(* PLC project PR_TT-1MasterSeq_Soft2.0_workflow_b380e4_PLC, SiemensToBackhoff Siemens TIA Portal → Beckhoff TwinCAT PLCopen Converter 2.2 *)
(* stored: creationDateTime 2026-10-12T09:25:48.748496, modificationDateTime 2026-10-12T09:25:48.748496 *)

FUNCTION_BLOCK PR_TT-1MasterSeq_Soft2.0_workflow_b380e4
VAR_INPUT
	iAllStationProcessOver : BOOL;
	iAutoRunning : BOOL;
	iHiPotTestOver_1 : BOOL;
	iHiPotTestOver_2 : BOOL;
	iHiPot_RTR_1 : BOOL;
	iHiPot_RTR_2 : BOOL;
	iIndexOver : BOOL;
	iIndex_RTR_Place1 : BOOL;
	iIndex_RTR_Place2 : BOOL;
	iOTS_Frm_Shuttle_1 : BOOL;
	iOTS_Frm_Shuttle_2 : BOOL;
	iOTS_Frm_TransferGantry : BOOL;
	iOperatorAck : BOOL;
	iPartPickOver : BOOL;
	iPartPickOver_1 : BOOL;
	iPartPickOver_2 : BOOL;
	iPartPlaceByTransferGantry : BOOL;
	iPartPlaceOver_IFGantry : BOOL;
	iPartPlaceOver_IndexPlace1 : BOOL;
	iPartPlaceOver_IndexPlace2 : BOOL;
	iPartPresent_IFGantry : BOOL;
	iPartPresent_Shuttle_1 : BOOL;
	iPartPresent_Shuttle_2 : BOOL;
	iPartPresent_TxGantry_1 : BOOL;
	iPartPresent_TxGantry_2 : BOOL;
	iRTR_Frm_TransferGantry_1 : BOOL;
	iRTR_Frm_TransferGantry_2 : BOOL;
	iReset_fault : BOOL;
	iShuttleReadyToReceive : BOOL;
	iSstMode : BOOL;
	iSstPB : BOOL;
END_VAR
VAR_OUTPUT
	qError : ARRAY[1..1] OF BOOL;
	qInfeedGantry_PickStart : BOOL;
	qInfeedGantry_PlaceStart : BOOL;
	qShuttle_1PickStart : BOOL;
	qShuttle_1PlaceStart : BOOL;
	qShuttle_2PickStart : BOOL;
	qShuttle_2PlaceStart : BOOL;
	qTransferGantry1_PickStart : BOOL;
	qTransferGantry1_PlaceStart : BOOL;
	qTransferGantry2_PickStart : BOOL;
	qTransferGantry2_PlaceStart : BOOL;
END_VAR
VAR
	c10_ChkPartStsAtSubStn_T1 : BOOL;
	c10_ChkPartStsAtSubStn_T2 : BOOL;
	c10_ChkPartStsAtSubStn_T3 : BOOL;
	c10_ChkPartStsAtSubStn_T4 : BOOL;
	c10_ChkPartStsAtSubStn_T5 : BOOL;
	c10_ChkPartStsAtSubStn_T6 : BOOL;
	c10_ChkPartStsAtSubStn_T7 : BOOL;
	c130_ChkPartPrsntStsShuttle2_T1 : BOOL;
	c130_ChkPartPrsntStsShuttle2_T2 : BOOL;
	c200_ChkPartPrsntTxGantry1_T1 : BOOL;
	c200_ChkPartPrsntTxGantry1_T2 : BOOL;
	c250_ChkPartPrsntTxGantry2_T1 : BOOL;
	c250_ChkPartPrsntTxGantry2_T2 : BOOL;
	c300_ChkPartPrsntIndexer_T1 : BOOL;
	c300_ChkPartPrsntIndexer_T2 : BOOL;
	c30_ChkPartStsIFGantry_T1 : BOOL;
	c30_ChkPartStsIFGantry_T2 : BOOL;
	c70_ChkPartPrsntStsShuttle1_T1 : BOOL;
	c70_ChkPartPrsntStsShuttle1_T2 : BOOL;
	StateNo : INT;
	s100_WtHiPotTestOver1 : BOOL;
	s100_WtHiPotTestOver1_T1 : BOOL;
	s10_ChkPartStsAtSubStn : BOOL;
	s10_ChkPartStsAtSubStn_T1 : BOOL;
	s10_ChkPartStsAtSubStn_T2 : BOOL;
	s10_ChkPartStsAtSubStn_T3 : BOOL;
	s10_ChkPartStsAtSubStn_T4 : BOOL;
	s10_ChkPartStsAtSubStn_T5 : BOOL;
	s10_ChkPartStsAtSubStn_T6 : BOOL;
	s10_ChkPartStsAtSubStn_T7 : BOOL;
	s110_WtTxGantryRTR1 : BOOL;
	s110_WtTxGantryRTR1_T1 : BOOL;
	s120_WtPartUnldOvrTxGantry1 : BOOL;
	s120_WtPartUnldOvrTxGantry1_T1 : BOOL;
	s130_ChkPartPrsntStsShuttle2 : BOOL;
	s130_ChkPartPrsntStsShuttle2_T1 : BOOL;
	s130_ChkPartPrsntStsShuttle2_T2 : BOOL;
	s140_WtIFGantryPlacePart2 : BOOL;
	s140_WtIFGantryPlacePart2_T1 : BOOL;
	s150_WtHiPotRdyRcvPart2 : BOOL;
	s150_WtHiPotRdyRcvPart2_T1 : BOOL;
	s160_WtHiPotTestOver2 : BOOL;
	s160_WtHiPotTestOver2_T1 : BOOL;
	s170_WtTxGantryRTR2 : BOOL;
	s170_WtTxGantryRTR2_T1 : BOOL;
	s190_WtPartUnldOvrTxGantry2 : BOOL;
	s190_WtPartUnldOvrTxGantry2_T1 : BOOL;
	s1_WtResetRel : BOOL;
	s1_WtResetRel_T1 : BOOL;
	s200_ChkPartPrsntTxGantry1 : BOOL;
	s200_ChkPartPrsntTxGantry1_T1 : BOOL;
	s200_ChkPartPrsntTxGantry1_T2 : BOOL;
	s20_WtOperatorAck : BOOL;
	s20_WtOperatorAck_T1 : BOOL;
	s210_WtShuttle1RdySendPal : BOOL;
	s210_WtShuttle1RdySendPal_T1 : BOOL;
	s220_WtPartPickTxGantry1 : BOOL;
	s220_WtPartPickTxGantry1_T1 : BOOL;
	s230_WtIndexRTRPlace1 : BOOL;
	s230_WtIndexRTRPlace1_T1 : BOOL;
	s240_WtPartPlaceOverIndexPlace1 : BOOL;
	s240_WtPartPlaceOverIndexPlace1_T1 : BOOL;
	s250_ChkPartPrsntTxGantry2 : BOOL;
	s250_ChkPartPrsntTxGantry2_T1 : BOOL;
	s250_ChkPartPrsntTxGantry2_T2 : BOOL;
	s260_WtShuttle2RdySendPal : BOOL;
	s260_WtShuttle2RdySendPal_T1 : BOOL;
	s270_WtPartPickTxGantry2 : BOOL;
	s270_WtPartPickTxGantry2_T1 : BOOL;
	s280_WtIndexRTRPlace2 : BOOL;
	s280_WtIndexRTRPlace2_T1 : BOOL;
	s290_WtPartPlaceOverIndexPlace2 : BOOL;
	s290_WtPartPlaceOverIndexPlace2_T1 : BOOL;
	s300_ChkPartPrsntIndexer : BOOL;
	s300_ChkPartPrsntIndexer_T1 : BOOL;
	s300_ChkPartPrsntIndexer_T2 : BOOL;
	s30_ChkPartStsIFGantry : BOOL;
	s30_ChkPartStsIFGantry_T1 : BOOL;
	s30_ChkPartStsIFGantry_T2 : BOOL;
	s310_WtOTSFrmTxGantry : BOOL;
	s310_WtOTSFrmTxGantry_T1 : BOOL;
	s320_WtPartPlaceByTxGantry : BOOL;
	s320_WtPartPlaceByTxGantry_T1 : BOOL;
	s330_WtAllStnProcessOver : BOOL;
	s330_WtAllStnProcessOver_T1 : BOOL;
	s340_WtIndexOver : BOOL;
	s340_WtIndexOver_T1 : BOOL;
	s40_WtPartPickOverIFGantry : BOOL;
	s40_WtPartPickOverIFGantry_T1 : BOOL;
	s50_WtShuttleRdyRcvPart : BOOL;
	s50_WtShuttleRdyRcvPart_T1 : BOOL;
	s60_WtPartPlaceByGantry : BOOL;
	s60_WtPartPlaceByGantry_T1 : BOOL;
	s70_ChkPartPrsntStsShuttle1 : BOOL;
	s70_ChkPartPrsntStsShuttle1_T1 : BOOL;
	s70_ChkPartPrsntStsShuttle1_T2 : BOOL;
	s80_WtIFGantryPlacePart : BOOL;
	s80_WtIFGantryPlacePart_T1 : BOOL;
	s90_WtHiPotRdyRcvPart1 : BOOL;
	s90_WtHiPotRdyRcvPart1_T1 : BOOL;
	sAbnormalCondition : BOOL;
	sIndexerSeq : BOOL;
	sInfeedGantry : BOOL;
	sPartAbsentAtAllStn : BOOL;
	sPartPrsntAtStn : BOOL;
	sShuttle_1Seq : BOOL;
	sShuttle_2Seq : BOOL;
	sSst : BOOL;
	sSstPulse : BOOL;
	sSstRise : R_TRIG;
	sStWtResetRel : BOOL;
	sStWtResetRel_T1 : BOOL;
	sTransferGantry_1Seq : BOOL;
	sTransferGantry_2Seq : BOOL;
END_VAR
VAR_TEMP
	tOne : BOOL;
END_VAR
  VAR  (* added by the conversion: wires and edge detectors of the diagram *)
    _w24 : BOOL;
    _w26 : BOOL;
    _w39 : BOOL;
    _w41 : BOOL;
    _w42 : BOOL;
    _w116 : BOOL;
    _w119 : BOOL;
    _w120 : BOOL;
    _w121 : BOOL;
    _w122 : BOOL;
    _w123 : BOOL;
    _w124 : BOOL;
    _w125 : BOOL;
    _w126 : BOOL;
    _w139 : BOOL;
    _w141 : BOOL;
    _w142 : BOOL;
    _w170 : BOOL;
    _w174 : BOOL;
    _w175 : BOOL;
    _w176 : BOOL;
    _w190 : BOOL;
    _w192 : BOOL;
    _w193 : BOOL;
    _w210 : BOOL;
    _w212 : BOOL;
    _w213 : BOOL;
    _w226 : BOOL;
    _w228 : BOOL;
    _w229 : BOOL;
    _w257 : BOOL;
    _w261 : BOOL;
    _w262 : BOOL;
    _w263 : BOOL;
    _w276 : BOOL;
    _w278 : BOOL;
    _w279 : BOOL;
    _w292 : BOOL;
    _w294 : BOOL;
    _w295 : BOOL;
    _w312 : BOOL;
    _w314 : BOOL;
    _w315 : BOOL;
    _w328 : BOOL;
    _w330 : BOOL;
    _w331 : BOOL;
    _w344 : BOOL;
    _w346 : BOOL;
    _w347 : BOOL;
    _w375 : BOOL;
    _w379 : BOOL;
    _w380 : BOOL;
    _w381 : BOOL;
    _w394 : BOOL;
    _w396 : BOOL;
    _w397 : BOOL;
    _w414 : BOOL;
    _w416 : BOOL;
    _w417 : BOOL;
    _w430 : BOOL;
    _w432 : BOOL;
    _w433 : BOOL;
    _w446 : BOOL;
    _w448 : BOOL;
    _w449 : BOOL;
    _w462 : BOOL;
    _w464 : BOOL;
    _w465 : BOOL;
    _w493 : BOOL;
    _w497 : BOOL;
    _w498 : BOOL;
    _w499 : BOOL;
    _w512 : BOOL;
    _w514 : BOOL;
    _w515 : BOOL;
    _w529 : BOOL;
    _w531 : BOOL;
    _w532 : BOOL;
    _w549 : BOOL;
    _w551 : BOOL;
    _w552 : BOOL;
    _w565 : BOOL;
    _w567 : BOOL;
    _w568 : BOOL;
    _w596 : BOOL;
    _w599 : BOOL;
    _w600 : BOOL;
    _w601 : BOOL;
    _w614 : BOOL;
    _w616 : BOOL;
    _w617 : BOOL;
    _w631 : BOOL;
    _w633 : BOOL;
    _w634 : BOOL;
    _w651 : BOOL;
    _w654 : BOOL;
    _w655 : BOOL;
    _w668 : BOOL;
    _w670 : BOOL;
    _w671 : BOOL;
    _w699 : BOOL;
    _w703 : BOOL;
    _w704 : BOOL;
    _w705 : BOOL;
    _w718 : BOOL;
    _w720 : BOOL;
    _w721 : BOOL;
    _w734 : BOOL;
    _w736 : BOOL;
    _w737 : BOOL;
    _w750 : BOOL;
    _w752 : BOOL;
    _w753 : BOOL;
    _w766 : BOOL;
    _w768 : BOOL;
    _w769 : BOOL;
  END_VAR

(* LD diagram, written out as Structured Text *)
(* Network 1 *)
(* Create Single Step Pulse bit *)
(* Create Single Step bit *)
(* Transition for STATE Num:0 Reset Released *)
(* STATE Num:0 Reset Released *)
(* Transition for STATE Num:1 Wait Reset Release *)
(* STATE Num:1 Wait Reset Release *)
(* Condition1 for STATE Num:10 Check Part Status at SubStation *)
(* Condition2 for STATE Num:10 Check Part Status at SubStation *)
(* Condition3 for STATE Num:10 Check Part Status at SubStation *)
(* Condition4 for STATE Num:10 Check Part Status at SubStation *)
(* Condition5 for STATE Num:10 Check Part Status at SubStation *)
(* Condition6 for STATE Num:10 Check Part Status at SubStation *)
(* Condition7 for STATE Num:10 Check Part Status at SubStation *)
(* Transition for STATE Num:10 Check Part Status at SubStation *)
(* STATE Num:10 Check Part Status at SubStation *)
(* Transition for STATE Num:20 Wait For Operator Ack *)
(* STATE Num:20 Wait For Operator Ack *)
(* Actions for STATE Num:20 Wait For Operator Ack *)
(* Condition1 for STATE Num:30 Check part Status at Infeed gantry *)
(* Condition2 for STATE Num:30 Check part Status at Infeed gantry *)
(* Transition for STATE Num:30 Check part Status at Infeed gantry *)
(* STATE Num:30 Check part Status at Infeed gantry *)
(* Transition for STATE Num:40 Wait For Part Pick Over By Infeed Gantry *)
(* STATE Num:40 Wait For Part Pick Over By Infeed Gantry *)
(* Actions for STATE Num:40 Wait For Part Pick Over By Infeed Gantry *)
(* Transition for STATE Num:50 Wait Shuttle Ready To Receive Part *)
(* STATE Num:50 Wait Shuttle Ready To Receive Part *)
(* Transition for STATE Num:60 Wait For Part Place By Gantry *)
(* STATE Num:60 Wait For Part Place By Gantry *)
(* Actions for STATE Num:60 Wait For Part Place By Gantry *)
(* Condition1 for STATE Num:70 Check Part Present Status At Shuttle-1 *)
(* Condition2 for STATE Num:70 Check Part Present Status At Shuttle-1 *)
(* Transition for STATE Num:70 Check Part Present Status At Shuttle-1 *)
(* STATE Num:70 Check Part Present Status At Shuttle-1 *)
(* Transition for STATE Num:80 Wait for Infeed Gantry Place Part *)
(* STATE Num:80 Wait for Infeed Gantry Place Part *)
(* Transition for STATE Num:90 Wait for HiPotReadyToReceivePart *)
(* STATE Num:90 Wait for HiPotReadyToReceivePart *)
(* Actions for STATE Num:90 Wait for HiPotReadyToReceivePart *)
(* Transition for STATE Num:100 Wait for HiPotTestOver_1 *)
(* STATE Num:100 Wait for HiPotTestOver_1 *)
(* Transition for STATE Num:110 Wait for Transfer Gantry Ready To Receive_1 *)
(* STATE Num:110 Wait for Transfer Gantry Ready To Receive_1 *)
(* Transition for STATE Num:120 Wait For part Unload Over from Transfer Gantry_1 *)
(* STATE Num:120 Wait For part Unload Over from Transfer Gantry_1 *)
(* Actions for STATE Num:120 Wait For part Unload Over from Transfer Gantry_1 *)
(* Condition1 for STATE Num:130 Check Part Present Status At Shuttle-2 *)
(* Condition2 for STATE Num:130 Check Part Present Status At Shuttle-2 *)
(* Transition for STATE Num:130 Check Part Present Status At Shuttle-2 *)
(* STATE Num:130 Check Part Present Status At Shuttle-2 *)
(* Transition for STATE Num:140 Wait for Infeed Gantry Place Part *)
(* STATE Num:140 Wait for Infeed Gantry Place Part *)
(* Actions for STATE Num:140 Wait for Infeed Gantry Place Part *)
(* Transition for STATE Num:150 Wait for HiPotReadyToReceivePart *)
(* STATE Num:150 Wait for HiPotReadyToReceivePart *)
(* Transition for STATE Num:160 Wait for HiPotTestOver_2 *)
(* STATE Num:160 Wait for HiPotTestOver_2 *)
(* Transition for STATE Num:170 Wait for Transfer Gantry Ready To Receive_2 *)
(* STATE Num:170 Wait for Transfer Gantry Ready To Receive_2 *)
(* Transition for STATE Num:190 Wait For part Unload Over from Transfer Gantry_2 *)
(* STATE Num:190 Wait For part Unload Over from Transfer Gantry_2 *)
(* Actions for STATE Num:190 Wait For part Unload Over from Transfer Gantry_2 *)
(* Condition1 for STATE Num:200 Check Part Present At Tranfer Gantry-1 *)
(* Condition2 for STATE Num:200 Check Part Present At Tranfer Gantry-1 *)
(* Transition for STATE Num:200 Check Part Present At Tranfer Gantry-1 *)
(* STATE Num:200 Check Part Present At Tranfer Gantry-1 *)
(* Transition for STATE Num:210 Wait for Shuttle-1 Ready to Send Pallet *)
(* STATE Num:210 Wait for Shuttle-1 Ready to Send Pallet *)
(* Transition for STATE Num:220 Wait for part Pick By Tranfer Gantry-1 *)
(* STATE Num:220 Wait for part Pick By Tranfer Gantry-1 *)
(* Actions for STATE Num:220 Wait for part Pick By Tranfer Gantry-1 *)
(* Transition for STATE Num:230 Wait for Indexer Ready to Receive_Place1 *)
(* STATE Num:230 Wait for Indexer Ready to Receive_Place1 *)
(* Transition for STATE Num:240 Wait for part Place Over Index Place1 *)
(* STATE Num:240 Wait for part Place Over Index Place1 *)
(* Actions for STATE Num:240 Wait for part Place Over Index Place1 *)
(* Condition1 for STATE Num:250 Check Part Present At Tranfer Gantry-2 *)
(* Condition2 for STATE Num:250 Check Part Present At Tranfer Gantry-2 *)
(* Transition for STATE Num:250 Check Part Present At Tranfer Gantry-2 *)
(* STATE Num:250 Check Part Present At Tranfer Gantry-2 *)
(* Transition for STATE Num:260 Wait for Shuttle-2 Ready to Send Pallet *)
(* STATE Num:260 Wait for Shuttle-2 Ready to Send Pallet *)
(* Transition for STATE Num:270 Wait for part Pick By Tranfer Gantry-2 *)
(* STATE Num:270 Wait for part Pick By Tranfer Gantry-2 *)
(* Actions for STATE Num:270 Wait for part Pick By Tranfer Gantry-2 *)
(* Transition for STATE Num:280 Wait for Indexer Ready to Receive_Place2 *)
(* STATE Num:280 Wait for Indexer Ready to Receive_Place2 *)
(* Transition for STATE Num:290 Wait for part Place Over Index Place2 *)
(* STATE Num:290 Wait for part Place Over Index Place2 *)
(* Actions for STATE Num:290 Wait for part Place Over Index Place2 *)
(* Condition1 for STATE Num:300 Check Part Present At Indexer *)
(* Condition2 for STATE Num:300 Check Part Present At Indexer *)
(* Transition for STATE Num:300 Check Part Present At Indexer *)
(* STATE Num:300 Check Part Present At Indexer *)
(* Transition for STATE Num:310 Wait for OTS From Transfer Gantry *)
(* STATE Num:310 Wait for OTS From Transfer Gantry *)
(* Transition for STATE Num:320 Wait for Part Place By Transfer Gantry *)
(* STATE Num:320 Wait for Part Place By Transfer Gantry *)
(* Transition for STATE Num:330 Wait All Station Process Over *)
(* STATE Num:330 Wait All Station Process Over *)
(* Transition for STATE Num:340 Wait for Index Over *)
(* STATE Num:340 Wait for Index Over *)
tOne := tOne OR NOT tOne;
sSstRise(CLK := iSstPB);
sSstPulse := sSstRise.Q;
sSst := iSstMode AND sSstPulse OR NOT iSstMode;
sStWtResetRel_T1 := sStWtResetRel AND iAutoRunning;
_w24 := sStWtResetRel;
_w26 := (_w24 OR NOT iAutoRunning) AND NOT sStWtResetRel_T1;
sStWtResetRel := _w26;
IF _w26 THEN StateNo := 0; END_IF;
s1_WtResetRel_T1 := s1_WtResetRel AND NOT sStWtResetRel AND sSst AND iAutoRunning;
_w39 := s1_WtResetRel;
_w41 := (_w39 OR sStWtResetRel_T1) AND NOT sStWtResetRel;
_w42 := _w41 AND NOT s1_WtResetRel_T1;
s1_WtResetRel := _w42;
IF _w42 THEN StateNo := 1; END_IF;
c10_ChkPartStsAtSubStn_T1 := sAbnormalCondition;
c10_ChkPartStsAtSubStn_T2 := sInfeedGantry;
c10_ChkPartStsAtSubStn_T3 := sShuttle_1Seq;
c10_ChkPartStsAtSubStn_T4 := sShuttle_2Seq;
c10_ChkPartStsAtSubStn_T5 := sTransferGantry_1Seq;
c10_ChkPartStsAtSubStn_T6 := sTransferGantry_2Seq;
c10_ChkPartStsAtSubStn_T7 := sIndexerSeq;
s10_ChkPartStsAtSubStn_T1 := s10_ChkPartStsAtSubStn AND NOT sStWtResetRel AND sSst AND c10_ChkPartStsAtSubStn_T1;
s10_ChkPartStsAtSubStn_T2 := s10_ChkPartStsAtSubStn AND NOT sStWtResetRel AND sSst AND NOT s10_ChkPartStsAtSubStn_T1 AND c10_ChkPartStsAtSubStn_T2;
s10_ChkPartStsAtSubStn_T3 := s10_ChkPartStsAtSubStn AND NOT sStWtResetRel AND sSst AND NOT s10_ChkPartStsAtSubStn_T1 AND NOT s10_ChkPartStsAtSubStn_T1 AND NOT s10_ChkPartStsAtSubStn_T2 AND c10_ChkPartStsAtSubStn_T3;
s10_ChkPartStsAtSubStn_T4 := s10_ChkPartStsAtSubStn AND NOT sStWtResetRel AND sSst AND NOT s10_ChkPartStsAtSubStn_T1 AND NOT s10_ChkPartStsAtSubStn_T1 AND NOT s10_ChkPartStsAtSubStn_T2 AND NOT s10_ChkPartStsAtSubStn_T1 AND NOT s10_ChkPartStsAtSubStn_T2 AND NOT s10_ChkPartStsAtSubStn_T3 AND c10_ChkPartStsAtSubStn_T4;
s10_ChkPartStsAtSubStn_T5 := s10_ChkPartStsAtSubStn AND NOT sStWtResetRel AND sSst AND NOT s10_ChkPartStsAtSubStn_T1 AND NOT s10_ChkPartStsAtSubStn_T1 AND NOT s10_ChkPartStsAtSubStn_T2 AND NOT s10_ChkPartStsAtSubStn_T1 AND NOT s10_ChkPartStsAtSubStn_T2 AND NOT s10_ChkPartStsAtSubStn_T3 AND NOT s10_ChkPartStsAtSubStn_T1 AND NOT s10_ChkPartStsAtSubStn_T2 AND NOT s10_ChkPartStsAtSubStn_T3 AND NOT s10_ChkPartStsAtSubStn_T4 AND c10_ChkPartStsAtSubStn_T5;
s10_ChkPartStsAtSubStn_T6 := s10_ChkPartStsAtSubStn AND NOT sStWtResetRel AND sSst AND NOT s10_ChkPartStsAtSubStn_T1 AND NOT s10_ChkPartStsAtSubStn_T1 AND NOT s10_ChkPartStsAtSubStn_T2 AND NOT s10_ChkPartStsAtSubStn_T1 AND NOT s10_ChkPartStsAtSubStn_T2 AND NOT s10_ChkPartStsAtSubStn_T3 AND NOT s10_ChkPartStsAtSubStn_T1 AND NOT s10_ChkPartStsAtSubStn_T2 AND NOT s10_ChkPartStsAtSubStn_T3 AND NOT s10_ChkPartStsAtSubStn_T4 AND NOT s10_ChkPartStsAtSubStn_T1 AND NOT s10_ChkPartStsAtSubStn_T2 AND NOT s10_ChkPartStsAtSubStn_T3 AND NOT s10_ChkPartStsAtSubStn_T4 AND NOT s10_ChkPartStsAtSubStn_T5 AND c10_ChkPartStsAtSubStn_T6;
s10_ChkPartStsAtSubStn_T7 := s10_ChkPartStsAtSubStn AND NOT sStWtResetRel AND sSst AND NOT s10_ChkPartStsAtSubStn_T1 AND NOT s10_ChkPartStsAtSubStn_T1 AND NOT s10_ChkPartStsAtSubStn_T2 AND NOT s10_ChkPartStsAtSubStn_T1 AND NOT s10_ChkPartStsAtSubStn_T2 AND NOT s10_ChkPartStsAtSubStn_T3 AND NOT s10_ChkPartStsAtSubStn_T1 AND NOT s10_ChkPartStsAtSubStn_T2 AND NOT s10_ChkPartStsAtSubStn_T3 AND NOT s10_ChkPartStsAtSubStn_T4 AND NOT s10_ChkPartStsAtSubStn_T1 AND NOT s10_ChkPartStsAtSubStn_T2 AND NOT s10_ChkPartStsAtSubStn_T3 AND NOT s10_ChkPartStsAtSubStn_T4 AND NOT s10_ChkPartStsAtSubStn_T5 AND NOT s10_ChkPartStsAtSubStn_T1 AND NOT s10_ChkPartStsAtSubStn_T2 AND NOT s10_ChkPartStsAtSubStn_T3 AND NOT s10_ChkPartStsAtSubStn_T4 AND NOT s10_ChkPartStsAtSubStn_T5 AND NOT s10_ChkPartStsAtSubStn_T6 AND c10_ChkPartStsAtSubStn_T7;
_w116 := s10_ChkPartStsAtSubStn;
_w119 := (_w116 OR s1_WtResetRel_T1 OR s20_WtOperatorAck_T1) AND NOT sStWtResetRel;
_w120 := _w119 AND NOT s10_ChkPartStsAtSubStn_T1;
_w121 := _w120 AND NOT s10_ChkPartStsAtSubStn_T2;
_w122 := _w121 AND NOT s10_ChkPartStsAtSubStn_T3;
_w123 := _w122 AND NOT s10_ChkPartStsAtSubStn_T4;
_w124 := _w123 AND NOT s10_ChkPartStsAtSubStn_T5;
_w125 := _w124 AND NOT s10_ChkPartStsAtSubStn_T6;
_w126 := _w125 AND NOT s10_ChkPartStsAtSubStn_T7;
s10_ChkPartStsAtSubStn := _w126;
IF _w126 THEN StateNo := 10; END_IF;
s20_WtOperatorAck_T1 := s20_WtOperatorAck AND NOT sStWtResetRel AND sSst AND iOperatorAck;
_w139 := s20_WtOperatorAck;
_w141 := (_w139 OR s10_ChkPartStsAtSubStn_T1) AND NOT sStWtResetRel;
_w142 := _w141 AND NOT s20_WtOperatorAck_T1;
s20_WtOperatorAck := _w142;
IF _w142 THEN StateNo := 20; END_IF;
qError[1] := s20_WtOperatorAck;
c30_ChkPartStsIFGantry_T1 := NOT iPartPresent_IFGantry;
c30_ChkPartStsIFGantry_T2 := iPartPresent_IFGantry;
s30_ChkPartStsIFGantry_T1 := s30_ChkPartStsIFGantry AND NOT sStWtResetRel AND sSst AND c30_ChkPartStsIFGantry_T1;
s30_ChkPartStsIFGantry_T2 := s30_ChkPartStsIFGantry AND NOT sStWtResetRel AND sSst AND NOT s30_ChkPartStsIFGantry_T1 AND c30_ChkPartStsIFGantry_T2;
_w170 := s30_ChkPartStsIFGantry;
_w174 := (_w170 OR s60_WtPartPlaceByGantry_T1 OR s10_ChkPartStsAtSubStn_T2 OR s40_WtPartPickOverIFGantry_T1) AND NOT sStWtResetRel;
_w175 := _w174 AND NOT s30_ChkPartStsIFGantry_T1;
_w176 := _w175 AND NOT s30_ChkPartStsIFGantry_T2;
s30_ChkPartStsIFGantry := _w176;
IF _w176 THEN StateNo := 30; END_IF;
s40_WtPartPickOverIFGantry_T1 := s40_WtPartPickOverIFGantry AND NOT sStWtResetRel AND sSst AND iPartPickOver AND iPartPresent_IFGantry;
_w190 := s40_WtPartPickOverIFGantry;
_w192 := (_w190 OR s30_ChkPartStsIFGantry_T1) AND NOT sStWtResetRel;
_w193 := _w192 AND NOT s40_WtPartPickOverIFGantry_T1;
s40_WtPartPickOverIFGantry := _w193;
IF _w193 THEN StateNo := 40; END_IF;
qInfeedGantry_PickStart := s40_WtPartPickOverIFGantry;
s50_WtShuttleRdyRcvPart_T1 := s50_WtShuttleRdyRcvPart AND NOT sStWtResetRel AND sSst AND iShuttleReadyToReceive;
_w210 := s50_WtShuttleRdyRcvPart;
_w212 := (_w210 OR s30_ChkPartStsIFGantry_T2) AND NOT sStWtResetRel;
_w213 := _w212 AND NOT s50_WtShuttleRdyRcvPart_T1;
s50_WtShuttleRdyRcvPart := _w213;
IF _w213 THEN StateNo := 50; END_IF;
s60_WtPartPlaceByGantry_T1 := s60_WtPartPlaceByGantry AND NOT sStWtResetRel AND sSst AND iPartPlaceOver_IFGantry;
_w226 := s60_WtPartPlaceByGantry;
_w228 := (_w226 OR s50_WtShuttleRdyRcvPart_T1) AND NOT sStWtResetRel;
_w229 := _w228 AND NOT s60_WtPartPlaceByGantry_T1;
s60_WtPartPlaceByGantry := _w229;
IF _w229 THEN StateNo := 60; END_IF;
qInfeedGantry_PlaceStart := s60_WtPartPlaceByGantry;
c70_ChkPartPrsntStsShuttle1_T1 := NOT iPartPresent_Shuttle_1;
c70_ChkPartPrsntStsShuttle1_T2 := iPartPresent_Shuttle_1;
s70_ChkPartPrsntStsShuttle1_T1 := s70_ChkPartPrsntStsShuttle1 AND NOT sStWtResetRel AND sSst AND c70_ChkPartPrsntStsShuttle1_T1;
s70_ChkPartPrsntStsShuttle1_T2 := s70_ChkPartPrsntStsShuttle1 AND NOT sStWtResetRel AND sSst AND NOT s70_ChkPartPrsntStsShuttle1_T1 AND c70_ChkPartPrsntStsShuttle1_T2;
_w257 := s70_ChkPartPrsntStsShuttle1;
_w261 := (_w257 OR s120_WtPartUnldOvrTxGantry1_T1 OR s10_ChkPartStsAtSubStn_T3 OR s80_WtIFGantryPlacePart_T1) AND NOT sStWtResetRel;
_w262 := _w261 AND NOT s70_ChkPartPrsntStsShuttle1_T1;
_w263 := _w262 AND NOT s70_ChkPartPrsntStsShuttle1_T2;
s70_ChkPartPrsntStsShuttle1 := _w263;
IF _w263 THEN StateNo := 70; END_IF;
s80_WtIFGantryPlacePart_T1 := s80_WtIFGantryPlacePart AND NOT sStWtResetRel AND sSst AND iPartPresent_Shuttle_1;
_w276 := s80_WtIFGantryPlacePart;
_w278 := (_w276 OR s70_ChkPartPrsntStsShuttle1_T1) AND NOT sStWtResetRel;
_w279 := _w278 AND NOT s80_WtIFGantryPlacePart_T1;
s80_WtIFGantryPlacePart := _w279;
IF _w279 THEN StateNo := 80; END_IF;
s90_WtHiPotRdyRcvPart1_T1 := s90_WtHiPotRdyRcvPart1 AND NOT sStWtResetRel AND sSst AND iHiPot_RTR_1;
_w292 := s90_WtHiPotRdyRcvPart1;
_w294 := (_w292 OR s70_ChkPartPrsntStsShuttle1_T2) AND NOT sStWtResetRel;
_w295 := _w294 AND NOT s90_WtHiPotRdyRcvPart1_T1;
s90_WtHiPotRdyRcvPart1 := _w295;
IF _w295 THEN StateNo := 90; END_IF;
qShuttle_1PlaceStart := s90_WtHiPotRdyRcvPart1;
s100_WtHiPotTestOver1_T1 := s100_WtHiPotTestOver1 AND NOT sStWtResetRel AND sSst AND iHiPotTestOver_1;
_w312 := s100_WtHiPotTestOver1;
_w314 := (_w312 OR s90_WtHiPotRdyRcvPart1_T1) AND NOT sStWtResetRel;
_w315 := _w314 AND NOT s100_WtHiPotTestOver1_T1;
s100_WtHiPotTestOver1 := _w315;
IF _w315 THEN StateNo := 100; END_IF;
s110_WtTxGantryRTR1_T1 := s110_WtTxGantryRTR1 AND NOT sStWtResetRel AND sSst AND iRTR_Frm_TransferGantry_1;
_w328 := s110_WtTxGantryRTR1;
_w330 := (_w328 OR s100_WtHiPotTestOver1_T1) AND NOT sStWtResetRel;
_w331 := _w330 AND NOT s110_WtTxGantryRTR1_T1;
s110_WtTxGantryRTR1 := _w331;
IF _w331 THEN StateNo := 110; END_IF;
s120_WtPartUnldOvrTxGantry1_T1 := s120_WtPartUnldOvrTxGantry1 AND NOT sStWtResetRel AND sSst AND NOT iPartPresent_Shuttle_1;
_w344 := s120_WtPartUnldOvrTxGantry1;
_w346 := (_w344 OR s110_WtTxGantryRTR1_T1) AND NOT sStWtResetRel;
_w347 := _w346 AND NOT s120_WtPartUnldOvrTxGantry1_T1;
s120_WtPartUnldOvrTxGantry1 := _w347;
IF _w347 THEN StateNo := 120; END_IF;
qShuttle_1PickStart := s120_WtPartUnldOvrTxGantry1;
c130_ChkPartPrsntStsShuttle2_T1 := NOT iPartPresent_Shuttle_2;
c130_ChkPartPrsntStsShuttle2_T2 := iPartPresent_Shuttle_2;
s130_ChkPartPrsntStsShuttle2_T1 := s130_ChkPartPrsntStsShuttle2 AND NOT sStWtResetRel AND sSst AND c130_ChkPartPrsntStsShuttle2_T1;
s130_ChkPartPrsntStsShuttle2_T2 := s130_ChkPartPrsntStsShuttle2 AND NOT sStWtResetRel AND sSst AND NOT s130_ChkPartPrsntStsShuttle2_T1 AND c130_ChkPartPrsntStsShuttle2_T2;
_w375 := s130_ChkPartPrsntStsShuttle2;
_w379 := (_w375 OR s190_WtPartUnldOvrTxGantry2_T1 OR s10_ChkPartStsAtSubStn_T4 OR s140_WtIFGantryPlacePart2_T1) AND NOT sStWtResetRel;
_w380 := _w379 AND NOT s130_ChkPartPrsntStsShuttle2_T1;
_w381 := _w380 AND NOT s130_ChkPartPrsntStsShuttle2_T2;
s130_ChkPartPrsntStsShuttle2 := _w381;
IF _w381 THEN StateNo := 130; END_IF;
s140_WtIFGantryPlacePart2_T1 := s140_WtIFGantryPlacePart2 AND NOT sStWtResetRel AND sSst AND iPartPresent_Shuttle_2;
_w394 := s140_WtIFGantryPlacePart2;
_w396 := (_w394 OR s130_ChkPartPrsntStsShuttle2_T1) AND NOT sStWtResetRel;
_w397 := _w396 AND NOT s140_WtIFGantryPlacePart2_T1;
s140_WtIFGantryPlacePart2 := _w397;
IF _w397 THEN StateNo := 140; END_IF;
qShuttle_2PlaceStart := s140_WtIFGantryPlacePart2;
s150_WtHiPotRdyRcvPart2_T1 := s150_WtHiPotRdyRcvPart2 AND NOT sStWtResetRel AND sSst AND iHiPot_RTR_2;
_w414 := s150_WtHiPotRdyRcvPart2;
_w416 := (_w414 OR s130_ChkPartPrsntStsShuttle2_T2) AND NOT sStWtResetRel;
_w417 := _w416 AND NOT s150_WtHiPotRdyRcvPart2_T1;
s150_WtHiPotRdyRcvPart2 := _w417;
IF _w417 THEN StateNo := 150; END_IF;
s160_WtHiPotTestOver2_T1 := s160_WtHiPotTestOver2 AND NOT sStWtResetRel AND sSst AND iHiPotTestOver_2;
_w430 := s160_WtHiPotTestOver2;
_w432 := (_w430 OR s150_WtHiPotRdyRcvPart2_T1) AND NOT sStWtResetRel;
_w433 := _w432 AND NOT s160_WtHiPotTestOver2_T1;
s160_WtHiPotTestOver2 := _w433;
IF _w433 THEN StateNo := 160; END_IF;
s170_WtTxGantryRTR2_T1 := s170_WtTxGantryRTR2 AND NOT sStWtResetRel AND sSst AND iRTR_Frm_TransferGantry_2;
_w446 := s170_WtTxGantryRTR2;
_w448 := (_w446 OR s160_WtHiPotTestOver2_T1) AND NOT sStWtResetRel;
_w449 := _w448 AND NOT s170_WtTxGantryRTR2_T1;
s170_WtTxGantryRTR2 := _w449;
IF _w449 THEN StateNo := 170; END_IF;
s190_WtPartUnldOvrTxGantry2_T1 := s190_WtPartUnldOvrTxGantry2 AND NOT sStWtResetRel AND sSst AND NOT iPartPresent_Shuttle_2;
_w462 := s190_WtPartUnldOvrTxGantry2;
_w464 := (_w462 OR s170_WtTxGantryRTR2_T1) AND NOT sStWtResetRel;
_w465 := _w464 AND NOT s190_WtPartUnldOvrTxGantry2_T1;
s190_WtPartUnldOvrTxGantry2 := _w465;
IF _w465 THEN StateNo := 190; END_IF;
qShuttle_2PickStart := s190_WtPartUnldOvrTxGantry2;
c200_ChkPartPrsntTxGantry1_T1 := NOT iPartPresent_TxGantry_1;
c200_ChkPartPrsntTxGantry1_T2 := iPartPresent_TxGantry_1;
s200_ChkPartPrsntTxGantry1_T1 := s200_ChkPartPrsntTxGantry1 AND NOT sStWtResetRel AND sSst AND c200_ChkPartPrsntTxGantry1_T1;
s200_ChkPartPrsntTxGantry1_T2 := s200_ChkPartPrsntTxGantry1 AND NOT sStWtResetRel AND sSst AND NOT s200_ChkPartPrsntTxGantry1_T1 AND c200_ChkPartPrsntTxGantry1_T2;
_w493 := s200_ChkPartPrsntTxGantry1;
_w497 := (_w493 OR s240_WtPartPlaceOverIndexPlace1_T1 OR s10_ChkPartStsAtSubStn_T5 OR s220_WtPartPickTxGantry1_T1) AND NOT sStWtResetRel;
_w498 := _w497 AND NOT s200_ChkPartPrsntTxGantry1_T1;
_w499 := _w498 AND NOT s200_ChkPartPrsntTxGantry1_T2;
s200_ChkPartPrsntTxGantry1 := _w499;
IF _w499 THEN StateNo := 200; END_IF;
s210_WtShuttle1RdySendPal_T1 := s210_WtShuttle1RdySendPal AND NOT sStWtResetRel AND sSst AND iOTS_Frm_Shuttle_1;
_w512 := s210_WtShuttle1RdySendPal;
_w514 := (_w512 OR s200_ChkPartPrsntTxGantry1_T1) AND NOT sStWtResetRel;
_w515 := _w514 AND NOT s210_WtShuttle1RdySendPal_T1;
s210_WtShuttle1RdySendPal := _w515;
IF _w515 THEN StateNo := 210; END_IF;
s220_WtPartPickTxGantry1_T1 := s220_WtPartPickTxGantry1 AND NOT sStWtResetRel AND sSst AND iPartPickOver_1 AND iPartPresent_TxGantry_1;
_w529 := s220_WtPartPickTxGantry1;
_w531 := (_w529 OR s210_WtShuttle1RdySendPal_T1) AND NOT sStWtResetRel;
_w532 := _w531 AND NOT s220_WtPartPickTxGantry1_T1;
s220_WtPartPickTxGantry1 := _w532;
IF _w532 THEN StateNo := 220; END_IF;
qTransferGantry1_PickStart := s220_WtPartPickTxGantry1;
s230_WtIndexRTRPlace1_T1 := s230_WtIndexRTRPlace1 AND NOT sStWtResetRel AND sSst AND iIndex_RTR_Place1;
_w549 := s230_WtIndexRTRPlace1;
_w551 := (_w549 OR s200_ChkPartPrsntTxGantry1_T2) AND NOT sStWtResetRel;
_w552 := _w551 AND NOT s230_WtIndexRTRPlace1_T1;
s230_WtIndexRTRPlace1 := _w552;
IF _w552 THEN StateNo := 230; END_IF;
s240_WtPartPlaceOverIndexPlace1_T1 := s240_WtPartPlaceOverIndexPlace1 AND NOT sStWtResetRel AND sSst AND iPartPlaceOver_IndexPlace1;
_w565 := s240_WtPartPlaceOverIndexPlace1;
_w567 := (_w565 OR s230_WtIndexRTRPlace1_T1) AND NOT sStWtResetRel;
_w568 := _w567 AND NOT s240_WtPartPlaceOverIndexPlace1_T1;
s240_WtPartPlaceOverIndexPlace1 := _w568;
IF _w568 THEN StateNo := 240; END_IF;
qTransferGantry1_PlaceStart := s240_WtPartPlaceOverIndexPlace1;
c250_ChkPartPrsntTxGantry2_T1 := NOT iPartPresent_TxGantry_2;
c250_ChkPartPrsntTxGantry2_T2 := iPartPresent_TxGantry_2;
s250_ChkPartPrsntTxGantry2_T1 := s250_ChkPartPrsntTxGantry2 AND NOT sStWtResetRel AND sSst AND c250_ChkPartPrsntTxGantry2_T1;
s250_ChkPartPrsntTxGantry2_T2 := s250_ChkPartPrsntTxGantry2 AND NOT sStWtResetRel AND sSst AND NOT s250_ChkPartPrsntTxGantry2_T1 AND c250_ChkPartPrsntTxGantry2_T2;
_w596 := s250_ChkPartPrsntTxGantry2;
_w599 := (_w596 OR s290_WtPartPlaceOverIndexPlace2_T1 OR s10_ChkPartStsAtSubStn_T6) AND NOT sStWtResetRel;
_w600 := _w599 AND NOT s250_ChkPartPrsntTxGantry2_T1;
_w601 := _w600 AND NOT s250_ChkPartPrsntTxGantry2_T2;
s250_ChkPartPrsntTxGantry2 := _w601;
IF _w601 THEN StateNo := 250; END_IF;
s260_WtShuttle2RdySendPal_T1 := s260_WtShuttle2RdySendPal AND NOT sStWtResetRel AND sSst AND iOTS_Frm_Shuttle_2;
_w614 := s260_WtShuttle2RdySendPal;
_w616 := (_w614 OR s250_ChkPartPrsntTxGantry2_T1) AND NOT sStWtResetRel;
_w617 := _w616 AND NOT s260_WtShuttle2RdySendPal_T1;
s260_WtShuttle2RdySendPal := _w617;
IF _w617 THEN StateNo := 260; END_IF;
s270_WtPartPickTxGantry2_T1 := s270_WtPartPickTxGantry2 AND NOT sStWtResetRel AND sSst AND iPartPickOver_2 AND iPartPresent_TxGantry_2;
_w631 := s270_WtPartPickTxGantry2;
_w633 := (_w631 OR s260_WtShuttle2RdySendPal_T1) AND NOT sStWtResetRel;
_w634 := _w633 AND NOT s270_WtPartPickTxGantry2_T1;
s270_WtPartPickTxGantry2 := _w634;
IF _w634 THEN StateNo := 270; END_IF;
qTransferGantry2_PickStart := s270_WtPartPickTxGantry2;
s280_WtIndexRTRPlace2_T1 := s280_WtIndexRTRPlace2 AND NOT sStWtResetRel AND sSst AND iIndex_RTR_Place2;
_w651 := s280_WtIndexRTRPlace2;
_w654 := (_w651 OR s270_WtPartPickTxGantry2_T1 OR s250_ChkPartPrsntTxGantry2_T2) AND NOT sStWtResetRel;
_w655 := _w654 AND NOT s280_WtIndexRTRPlace2_T1;
s280_WtIndexRTRPlace2 := _w655;
IF _w655 THEN StateNo := 280; END_IF;
s290_WtPartPlaceOverIndexPlace2_T1 := s290_WtPartPlaceOverIndexPlace2 AND NOT sStWtResetRel AND sSst AND iPartPlaceOver_IndexPlace2;
_w668 := s290_WtPartPlaceOverIndexPlace2;
_w670 := (_w668 OR s280_WtIndexRTRPlace2_T1) AND NOT sStWtResetRel;
_w671 := _w670 AND NOT s290_WtPartPlaceOverIndexPlace2_T1;
s290_WtPartPlaceOverIndexPlace2 := _w671;
IF _w671 THEN StateNo := 290; END_IF;
qTransferGantry2_PlaceStart := s290_WtPartPlaceOverIndexPlace2;
c300_ChkPartPrsntIndexer_T1 := sPartAbsentAtAllStn;
c300_ChkPartPrsntIndexer_T2 := sPartPrsntAtStn;
s300_ChkPartPrsntIndexer_T1 := s300_ChkPartPrsntIndexer AND NOT sStWtResetRel AND sSst AND c300_ChkPartPrsntIndexer_T1;
s300_ChkPartPrsntIndexer_T2 := s300_ChkPartPrsntIndexer AND NOT sStWtResetRel AND sSst AND NOT s300_ChkPartPrsntIndexer_T1 AND c300_ChkPartPrsntIndexer_T2;
_w699 := s300_ChkPartPrsntIndexer;
_w703 := (_w699 OR s340_WtIndexOver_T1 OR s10_ChkPartStsAtSubStn_T7 OR s320_WtPartPlaceByTxGantry_T1) AND NOT sStWtResetRel;
_w704 := _w703 AND NOT s300_ChkPartPrsntIndexer_T1;
_w705 := _w704 AND NOT s300_ChkPartPrsntIndexer_T2;
s300_ChkPartPrsntIndexer := _w705;
IF _w705 THEN StateNo := 300; END_IF;
s310_WtOTSFrmTxGantry_T1 := s310_WtOTSFrmTxGantry AND NOT sStWtResetRel AND sSst AND iOTS_Frm_TransferGantry;
_w718 := s310_WtOTSFrmTxGantry;
_w720 := (_w718 OR s300_ChkPartPrsntIndexer_T1) AND NOT sStWtResetRel;
_w721 := _w720 AND NOT s310_WtOTSFrmTxGantry_T1;
s310_WtOTSFrmTxGantry := _w721;
IF _w721 THEN StateNo := 310; END_IF;
s320_WtPartPlaceByTxGantry_T1 := s320_WtPartPlaceByTxGantry AND NOT sStWtResetRel AND sSst AND iPartPlaceByTransferGantry;
_w734 := s320_WtPartPlaceByTxGantry;
_w736 := (_w734 OR s310_WtOTSFrmTxGantry_T1) AND NOT sStWtResetRel;
_w737 := _w736 AND NOT s320_WtPartPlaceByTxGantry_T1;
s320_WtPartPlaceByTxGantry := _w737;
IF _w737 THEN StateNo := 320; END_IF;
s330_WtAllStnProcessOver_T1 := s330_WtAllStnProcessOver AND NOT sStWtResetRel AND sSst AND iAllStationProcessOver;
_w750 := s330_WtAllStnProcessOver;
_w752 := (_w750 OR s300_ChkPartPrsntIndexer_T2) AND NOT sStWtResetRel;
_w753 := _w752 AND NOT s330_WtAllStnProcessOver_T1;
s330_WtAllStnProcessOver := _w753;
IF _w753 THEN StateNo := 330; END_IF;
s340_WtIndexOver_T1 := s340_WtIndexOver AND NOT sStWtResetRel AND sSst AND iIndexOver;
_w766 := s340_WtIndexOver;
_w768 := (_w766 OR s330_WtAllStnProcessOver_T1) AND NOT sStWtResetRel;
_w769 := _w768 AND NOT s340_WtIndexOver_T1;
s340_WtIndexOver := _w769;
IF _w769 THEN StateNo := 340; END_IF;
END_FUNCTION_BLOCK
